// Mitsubishi GX Works2 project: B_v6_split   PLC: Q03UDE

PROGRAM COMMON
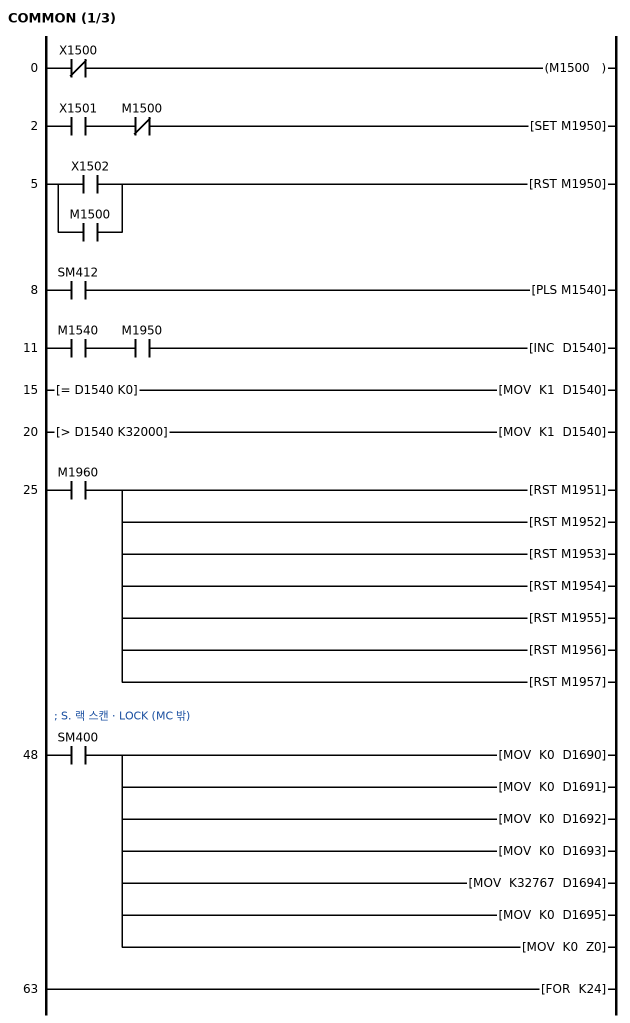
0     LDI     X1500
      OUT     M1500
2     LD      X1501
      ANI     M1500
      SET     M1950
5     LD      X1502
      OR      M1500
      RST     M1950
8     LD      SM412
      PLS     M1540
11    LD      M1540
      AND     M1950
      INC     D1540
15    LD=     D1540 K0
      MOV     K1 D1540
20    LD>     D1540 K32000
      MOV     K1 D1540
25    LD      M1960
      RST     M1951
      RST     M1952
      RST     M1953
      RST     M1954
      RST     M1955
      RST     M1956
      RST     M1957
; S. 랙 스캔 · LOCK (MC 밖)
48    LD      SM400
      MOV     K0 D1690
      MOV     K0 D1691
      MOV     K0 D1692
      MOV     K0 D1693
      MOV     K32767 D1694
      MOV     K0 D1695
      MOV     K0 Z0
63    FOR     K24
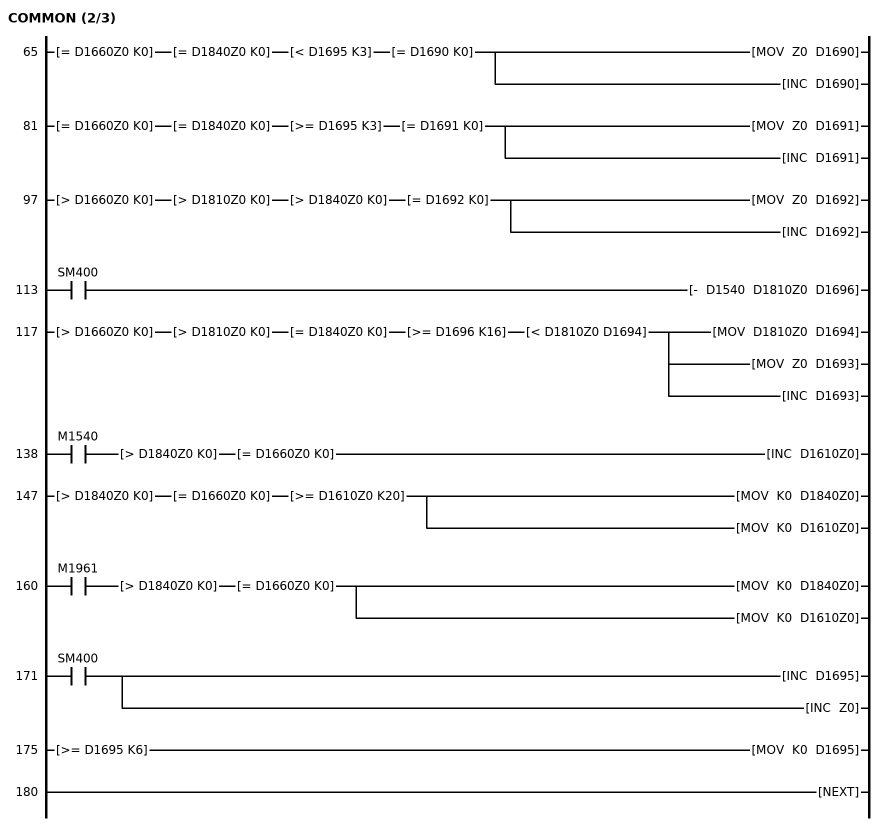
65    LD=     D1660Z0 K0
      AND=    D1840Z0 K0
      AND<    D1695 K3
      AND=    D1690 K0
      MOV     Z0 D1690
      INC     D1690
81    LD=     D1660Z0 K0
      AND=    D1840Z0 K0
      AND>=   D1695 K3
      AND=    D1691 K0
      MOV     Z0 D1691
      INC     D1691
97    LD>     D1660Z0 K0
      AND>    D1810Z0 K0
      AND>    D1840Z0 K0
      AND=    D1692 K0
      MOV     Z0 D1692
      INC     D1692
113   LD      SM400
      -       D1540 D1810Z0 D1696
117   LD>     D1660Z0 K0
      AND>    D1810Z0 K0
      AND=    D1840Z0 K0
      AND>=   D1696 K16
      AND<    D1810Z0 D1694
      MOV     D1810Z0 D1694
      MOV     Z0 D1693
      INC     D1693
138   LD      M1540
      AND>    D1840Z0 K0
      AND=    D1660Z0 K0
      INC     D1610Z0
147   LD>     D1840Z0 K0
      AND=    D1660Z0 K0
      AND>=   D1610Z0 K20
      MOV     K0 D1840Z0
      MOV     K0 D1610Z0
160   LD      M1961
      AND>    D1840Z0 K0
      AND=    D1660Z0 K0
      MOV     K0 D1840Z0
      MOV     K0 D1610Z0
171   LD      SM400
      INC     D1695
      INC     Z0
175   LD>=    D1695 K6
      MOV     K0 D1695
180   NEXT
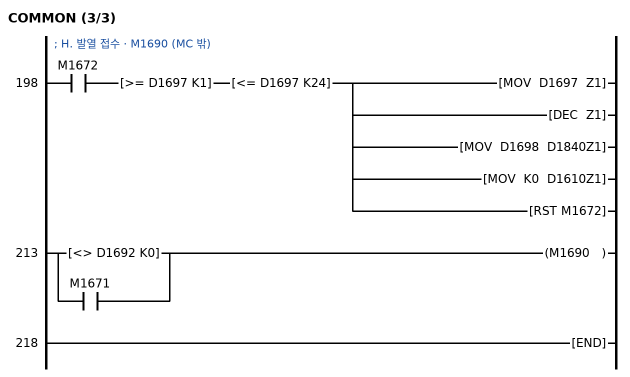
; H. 발열 접수 · M1690 (MC 밖)
198   LD      M1672
      AND>=   D1697 K1
      AND<=   D1697 K24
      MOV     D1697 Z1
      DEC     Z1
      MOV     D1698 D1840Z1
      MOV     K0 D1610Z1
      RST     M1672
213   LD<>    D1692 K0
      OR      M1671
      OUT     M1690
218   END
END_PROGRAM

PROGRAM RFID
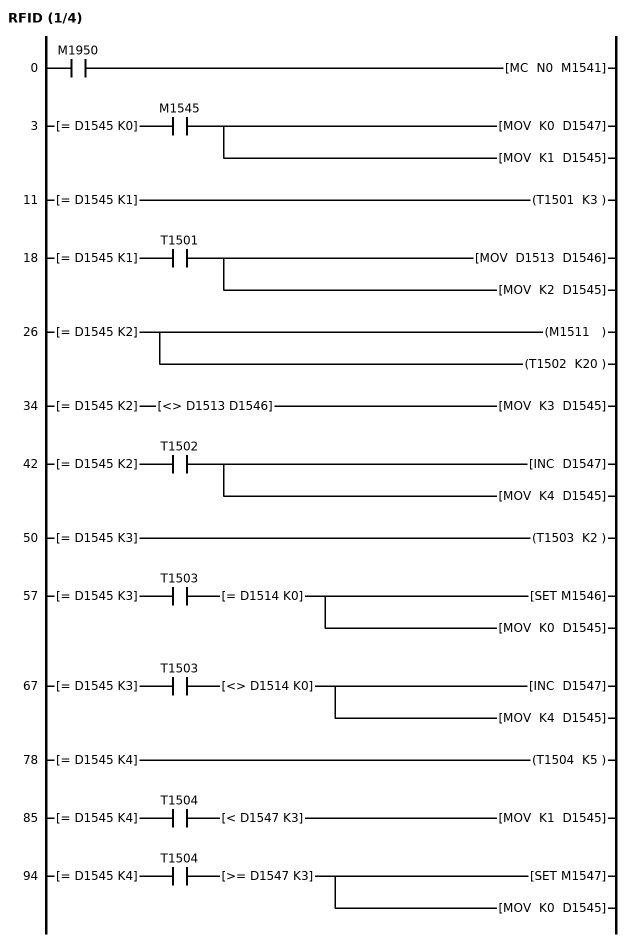
0     LD      M1950
      MC      N0 M1541
3     LD=     D1545 K0
      AND     M1545
      MOV     K0 D1547
      MOV     K1 D1545
11    LD=     D1545 K1
      OUT     T1501 K3
18    LD=     D1545 K1
      AND     T1501
      MOV     D1513 D1546
      MOV     K2 D1545
26    LD=     D1545 K2
      OUT     M1511
      OUT     T1502 K20
34    LD=     D1545 K2
      AND<>   D1513 D1546
      MOV     K3 D1545
42    LD=     D1545 K2
      AND     T1502
      INC     D1547
      MOV     K4 D1545
50    LD=     D1545 K3
      OUT     T1503 K2
57    LD=     D1545 K3
      AND     T1503
      AND=    D1514 K0
      SET     M1546
      MOV     K0 D1545
67    LD=     D1545 K3
      AND     T1503
      AND<>   D1514 K0
      INC     D1547
      MOV     K4 D1545
78    LD=     D1545 K4
      OUT     T1504 K5
85    LD=     D1545 K4
      AND     T1504
      AND<    D1547 K3
      MOV     K1 D1545
94    LD=     D1545 K4
      AND     T1504
      AND>=   D1547 K3
      SET     M1547
      MOV     K0 D1545
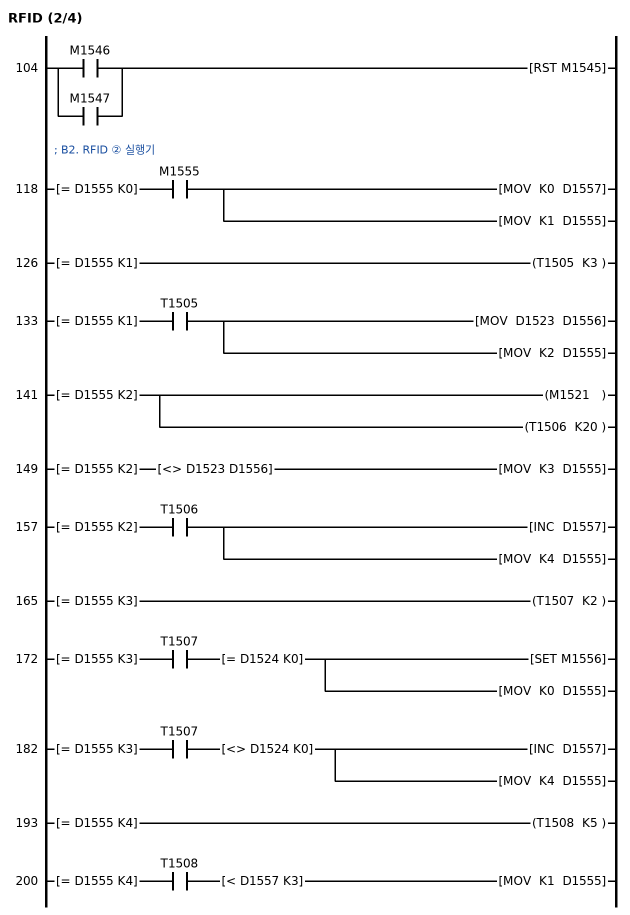
104   LD      M1546
      OR      M1547
      RST     M1545
; B2. RFID ② 실행기
118   LD=     D1555 K0
      AND     M1555
      MOV     K0 D1557
      MOV     K1 D1555
126   LD=     D1555 K1
      OUT     T1505 K3
133   LD=     D1555 K1
      AND     T1505
      MOV     D1523 D1556
      MOV     K2 D1555
141   LD=     D1555 K2
      OUT     M1521
      OUT     T1506 K20
149   LD=     D1555 K2
      AND<>   D1523 D1556
      MOV     K3 D1555
157   LD=     D1555 K2
      AND     T1506
      INC     D1557
      MOV     K4 D1555
165   LD=     D1555 K3
      OUT     T1507 K2
172   LD=     D1555 K3
      AND     T1507
      AND=    D1524 K0
      SET     M1556
      MOV     K0 D1555
182   LD=     D1555 K3
      AND     T1507
      AND<>   D1524 K0
      INC     D1557
      MOV     K4 D1555
193   LD=     D1555 K4
      OUT     T1508 K5
200   LD=     D1555 K4
      AND     T1508
      AND<    D1557 K3
      MOV     K1 D1555
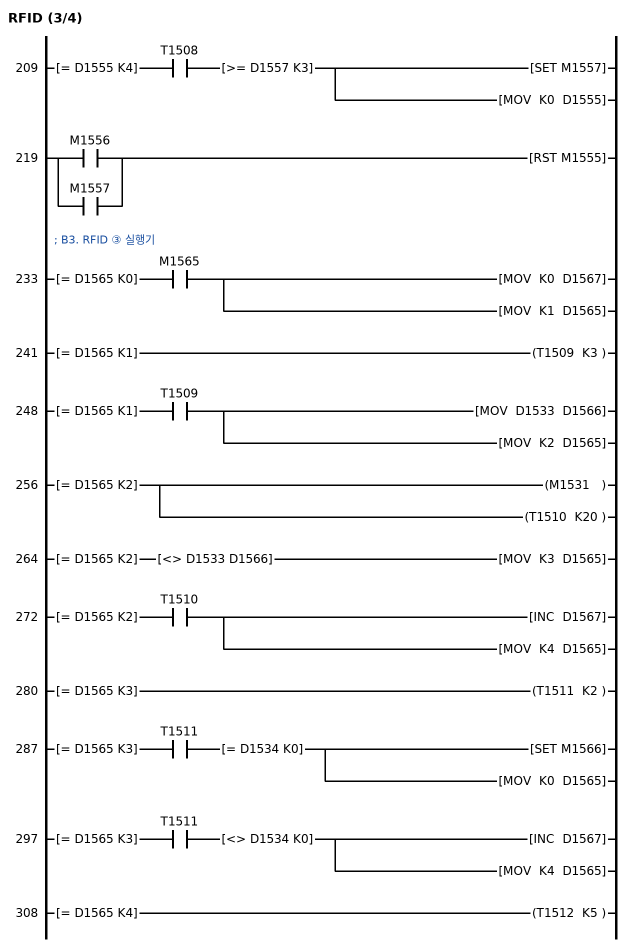
209   LD=     D1555 K4
      AND     T1508
      AND>=   D1557 K3
      SET     M1557
      MOV     K0 D1555
219   LD      M1556
      OR      M1557
      RST     M1555
; B3. RFID ③ 실행기
233   LD=     D1565 K0
      AND     M1565
      MOV     K0 D1567
      MOV     K1 D1565
241   LD=     D1565 K1
      OUT     T1509 K3
248   LD=     D1565 K1
      AND     T1509
      MOV     D1533 D1566
      MOV     K2 D1565
256   LD=     D1565 K2
      OUT     M1531
      OUT     T1510 K20
264   LD=     D1565 K2
      AND<>   D1533 D1566
      MOV     K3 D1565
272   LD=     D1565 K2
      AND     T1510
      INC     D1567
      MOV     K4 D1565
280   LD=     D1565 K3
      OUT     T1511 K2
287   LD=     D1565 K3
      AND     T1511
      AND=    D1534 K0
      SET     M1566
      MOV     K0 D1565
297   LD=     D1565 K3
      AND     T1511
      AND<>   D1534 K0
      INC     D1567
      MOV     K4 D1565
308   LD=     D1565 K4
      OUT     T1512 K5
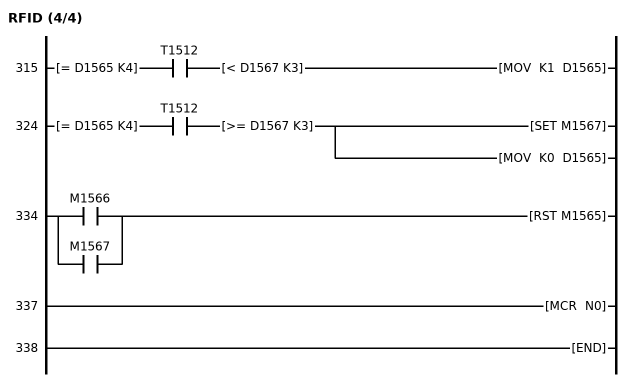
315   LD=     D1565 K4
      AND     T1512
      AND<    D1567 K3
      MOV     K1 D1565
324   LD=     D1565 K4
      AND     T1512
      AND>=   D1567 K3
      SET     M1567
      MOV     K0 D1565
334   LD      M1566
      OR      M1567
      RST     M1565
337   MCR     N0
338   END
END_PROGRAM

PROGRAM INFEED
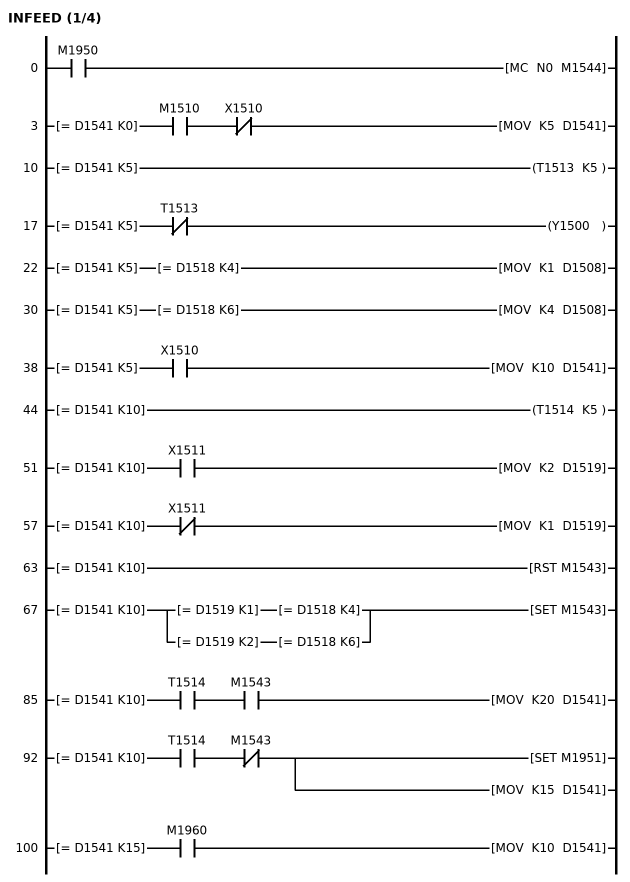
0     LD      M1950
      MC      N0 M1544
3     LD=     D1541 K0
      AND     M1510
      ANI     X1510
      MOV     K5 D1541
10    LD=     D1541 K5
      OUT     T1513 K5
17    LD=     D1541 K5
      ANI     T1513
      OUT     Y1500
22    LD=     D1541 K5
      AND=    D1518 K4
      MOV     K1 D1508
30    LD=     D1541 K5
      AND=    D1518 K6
      MOV     K4 D1508
38    LD=     D1541 K5
      AND     X1510
      MOV     K10 D1541
44    LD=     D1541 K10
      OUT     T1514 K5
51    LD=     D1541 K10
      AND     X1511
      MOV     K2 D1519
57    LD=     D1541 K10
      ANI     X1511
      MOV     K1 D1519
63    LD=     D1541 K10
      RST     M1543
67    LD=     D1541 K10
      LD=     D1519 K1
      AND=    D1518 K4
      LD=     D1519 K2
      AND=    D1518 K6
      ORB
      ANB
      SET     M1543
85    LD=     D1541 K10
      AND     T1514
      AND     M1543
      MOV     K20 D1541
92    LD=     D1541 K10
      AND     T1514
      ANI     M1543
      SET     M1951
      MOV     K15 D1541
100   LD=     D1541 K15
      AND     M1960
      MOV     K10 D1541
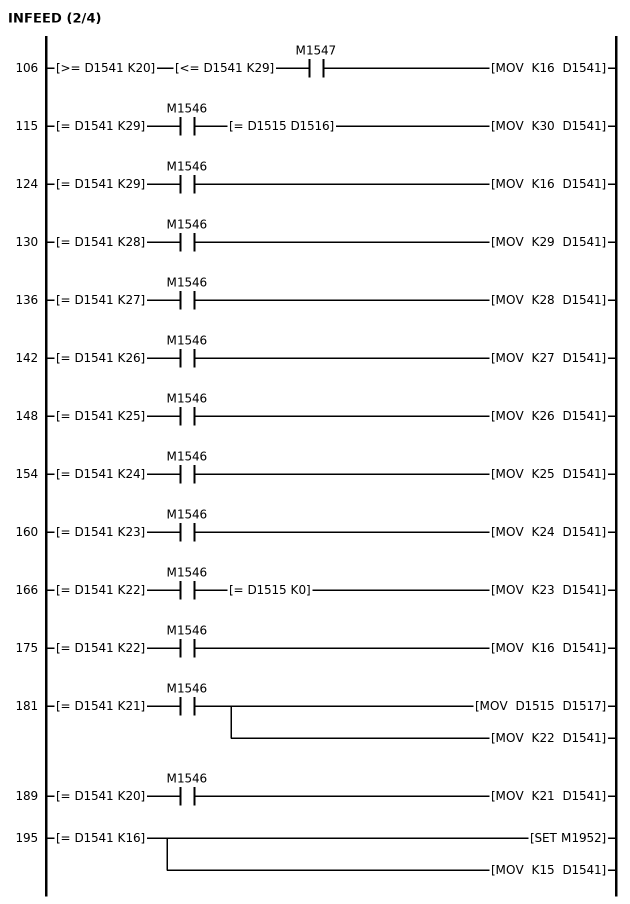
106   LD>=    D1541 K20
      AND<=   D1541 K29
      AND     M1547
      MOV     K16 D1541
115   LD=     D1541 K29
      AND     M1546
      AND=    D1515 D1516
      MOV     K30 D1541
124   LD=     D1541 K29
      AND     M1546
      MOV     K16 D1541
130   LD=     D1541 K28
      AND     M1546
      MOV     K29 D1541
136   LD=     D1541 K27
      AND     M1546
      MOV     K28 D1541
142   LD=     D1541 K26
      AND     M1546
      MOV     K27 D1541
148   LD=     D1541 K25
      AND     M1546
      MOV     K26 D1541
154   LD=     D1541 K24
      AND     M1546
      MOV     K25 D1541
160   LD=     D1541 K23
      AND     M1546
      MOV     K24 D1541
166   LD=     D1541 K22
      AND     M1546
      AND=    D1515 K0
      MOV     K23 D1541
175   LD=     D1541 K22
      AND     M1546
      MOV     K16 D1541
181   LD=     D1541 K21
      AND     M1546
      MOV     D1515 D1517
      MOV     K22 D1541
189   LD=     D1541 K20
      AND     M1546
      MOV     K21 D1541
195   LD=     D1541 K16
      SET     M1952
      MOV     K15 D1541
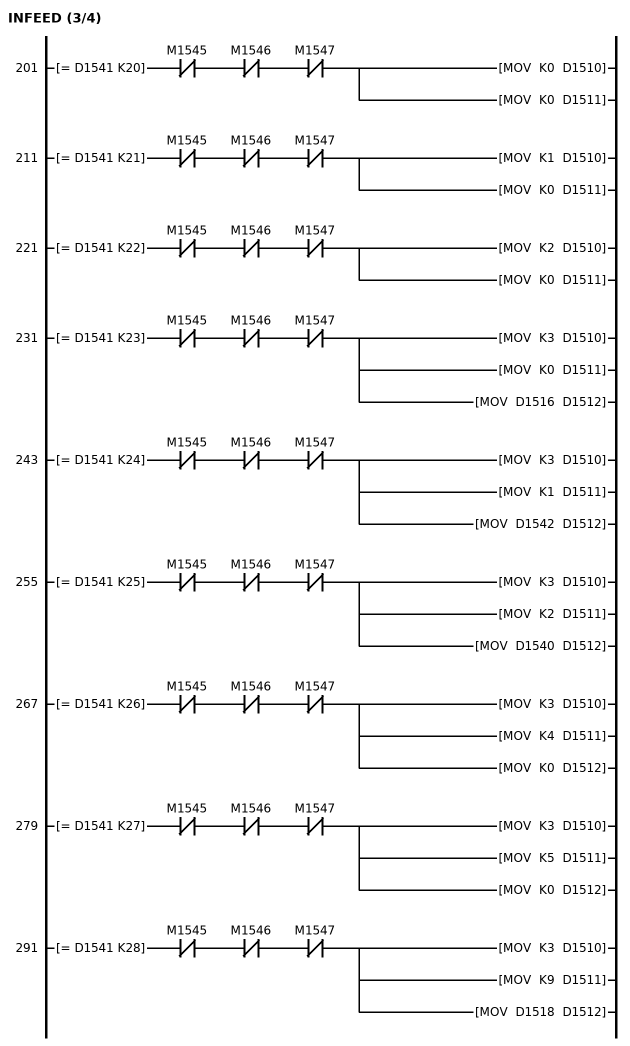
201   LD=     D1541 K20
      ANI     M1545
      ANI     M1546
      ANI     M1547
      MOV     K0 D1510
      MOV     K0 D1511
211   LD=     D1541 K21
      ANI     M1545
      ANI     M1546
      ANI     M1547
      MOV     K1 D1510
      MOV     K0 D1511
221   LD=     D1541 K22
      ANI     M1545
      ANI     M1546
      ANI     M1547
      MOV     K2 D1510
      MOV     K0 D1511
231   LD=     D1541 K23
      ANI     M1545
      ANI     M1546
      ANI     M1547
      MOV     K3 D1510
      MOV     K0 D1511
      MOV     D1516 D1512
243   LD=     D1541 K24
      ANI     M1545
      ANI     M1546
      ANI     M1547
      MOV     K3 D1510
      MOV     K1 D1511
      MOV     D1542 D1512
255   LD=     D1541 K25
      ANI     M1545
      ANI     M1546
      ANI     M1547
      MOV     K3 D1510
      MOV     K2 D1511
      MOV     D1540 D1512
267   LD=     D1541 K26
      ANI     M1545
      ANI     M1546
      ANI     M1547
      MOV     K3 D1510
      MOV     K4 D1511
      MOV     K0 D1512
279   LD=     D1541 K27
      ANI     M1545
      ANI     M1546
      ANI     M1547
      MOV     K3 D1510
      MOV     K5 D1511
      MOV     K0 D1512
291   LD=     D1541 K28
      ANI     M1545
      ANI     M1546
      ANI     M1547
      MOV     K3 D1510
      MOV     K9 D1511
      MOV     D1518 D1512
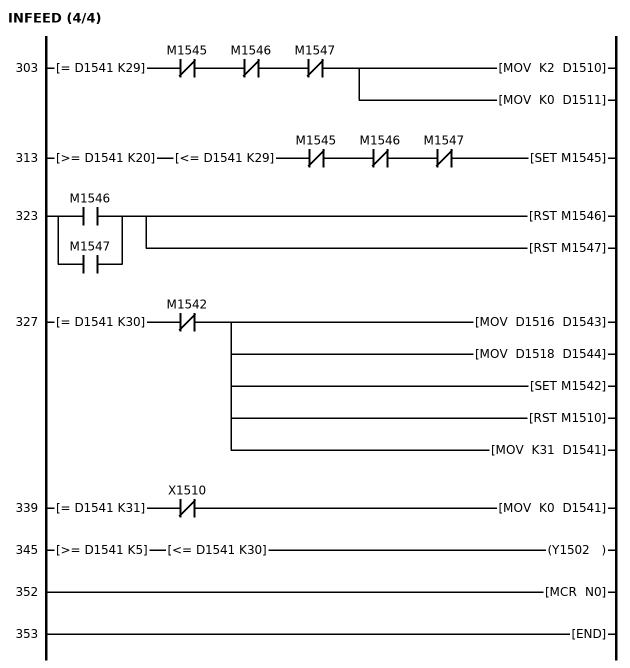
303   LD=     D1541 K29
      ANI     M1545
      ANI     M1546
      ANI     M1547
      MOV     K2 D1510
      MOV     K0 D1511
313   LD>=    D1541 K20
      AND<=   D1541 K29
      ANI     M1545
      ANI     M1546
      ANI     M1547
      SET     M1545
323   LD      M1546
      OR      M1547
      RST     M1546
      RST     M1547
327   LD=     D1541 K30
      ANI     M1542
      MOV     D1516 D1543
      MOV     D1518 D1544
      SET     M1542
      RST     M1510
      MOV     K31 D1541
339   LD=     D1541 K31
      ANI     X1510
      MOV     K0 D1541
345   LD>=    D1541 K5
      AND<=   D1541 K30
      OUT     Y1502
352   MCR     N0
353   END
END_PROGRAM

PROGRAM CRANE
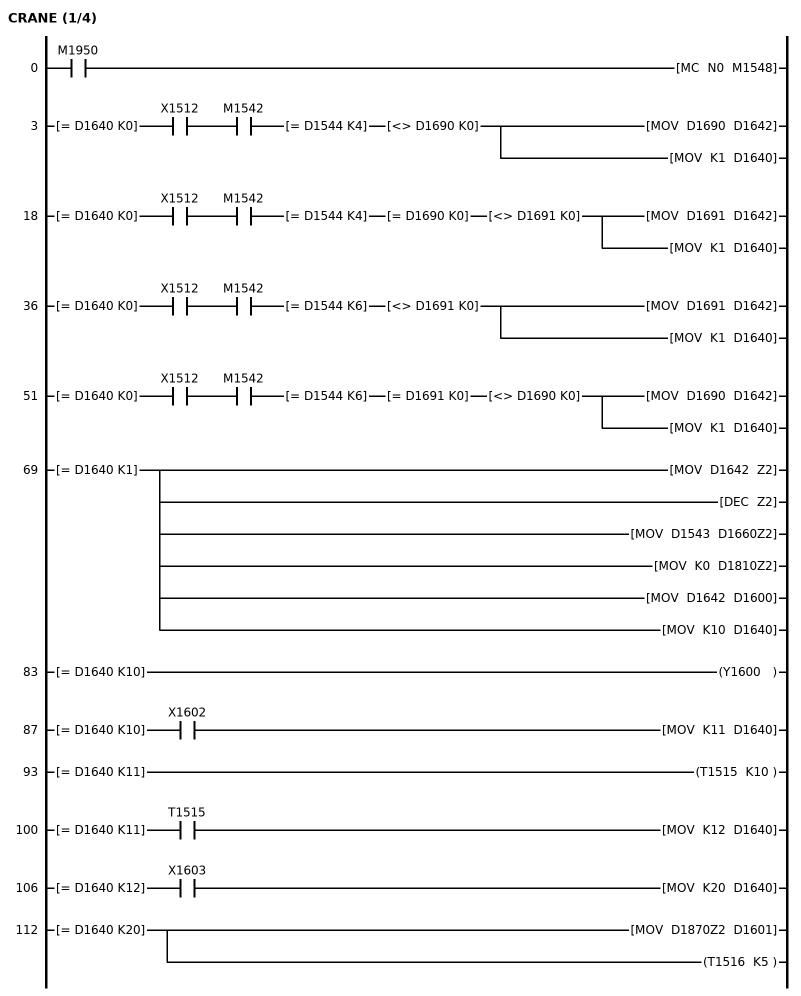
0     LD      M1950
      MC      N0 M1548
3     LD=     D1640 K0
      AND     X1512
      AND     M1542
      AND=    D1544 K4
      AND<>   D1690 K0
      MOV     D1690 D1642
      MOV     K1 D1640
18    LD=     D1640 K0
      AND     X1512
      AND     M1542
      AND=    D1544 K4
      AND=    D1690 K0
      AND<>   D1691 K0
      MOV     D1691 D1642
      MOV     K1 D1640
36    LD=     D1640 K0
      AND     X1512
      AND     M1542
      AND=    D1544 K6
      AND<>   D1691 K0
      MOV     D1691 D1642
      MOV     K1 D1640
51    LD=     D1640 K0
      AND     X1512
      AND     M1542
      AND=    D1544 K6
      AND=    D1691 K0
      AND<>   D1690 K0
      MOV     D1690 D1642
      MOV     K1 D1640
69    LD=     D1640 K1
      MOV     D1642 Z2
      DEC     Z2
      MOV     D1543 D1660Z2
      MOV     K0 D1810Z2
      MOV     D1642 D1600
      MOV     K10 D1640
83    LD=     D1640 K10
      OUT     Y1600
87    LD=     D1640 K10
      AND     X1602
      MOV     K11 D1640
93    LD=     D1640 K11
      OUT     T1515 K10
100   LD=     D1640 K11
      AND     T1515
      MOV     K12 D1640
106   LD=     D1640 K12
      AND     X1603
      MOV     K20 D1640
112   LD=     D1640 K20
      MOV     D1870Z2 D1601
      OUT     T1516 K5
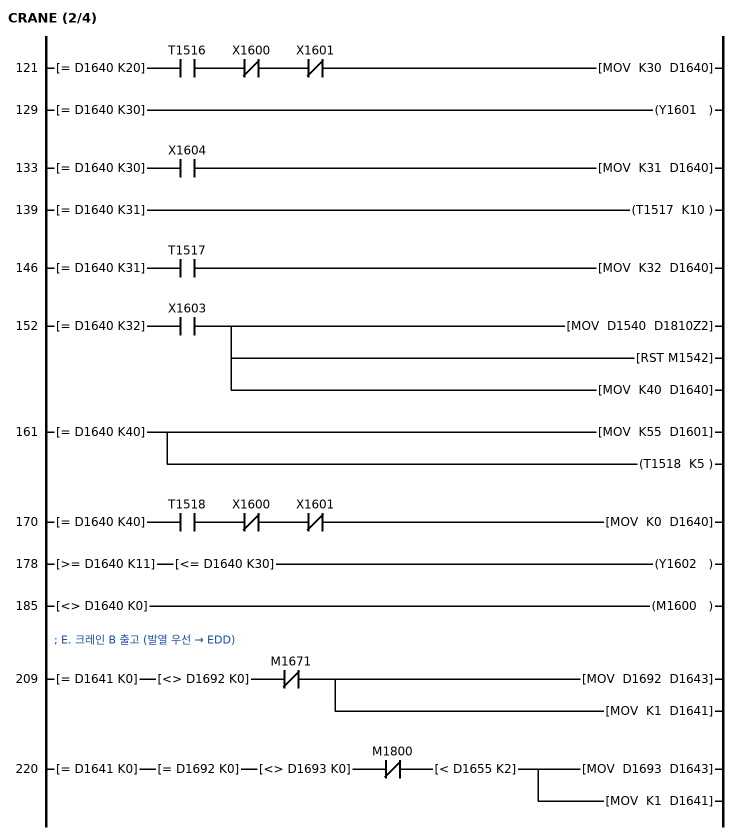
121   LD=     D1640 K20
      AND     T1516
      ANI     X1600
      ANI     X1601
      MOV     K30 D1640
129   LD=     D1640 K30
      OUT     Y1601
133   LD=     D1640 K30
      AND     X1604
      MOV     K31 D1640
139   LD=     D1640 K31
      OUT     T1517 K10
146   LD=     D1640 K31
      AND     T1517
      MOV     K32 D1640
152   LD=     D1640 K32
      AND     X1603
      MOV     D1540 D1810Z2
      RST     M1542
      MOV     K40 D1640
161   LD=     D1640 K40
      MOV     K55 D1601
      OUT     T1518 K5
170   LD=     D1640 K40
      AND     T1518
      ANI     X1600
      ANI     X1601
      MOV     K0 D1640
178   LD>=    D1640 K11
      AND<=   D1640 K30
      OUT     Y1602
185   LD<>    D1640 K0
      OUT     M1600
; E. 크레인 B 출고 (발열 우선 → EDD)
209   LD=     D1641 K0
      AND<>   D1692 K0
      ANI     M1671
      MOV     D1692 D1643
      MOV     K1 D1641
220   LD=     D1641 K0
      AND=    D1692 K0
      AND<>   D1693 K0
      ANI     M1800
      AND<    D1655 K2
      MOV     D1693 D1643
      MOV     K1 D1641
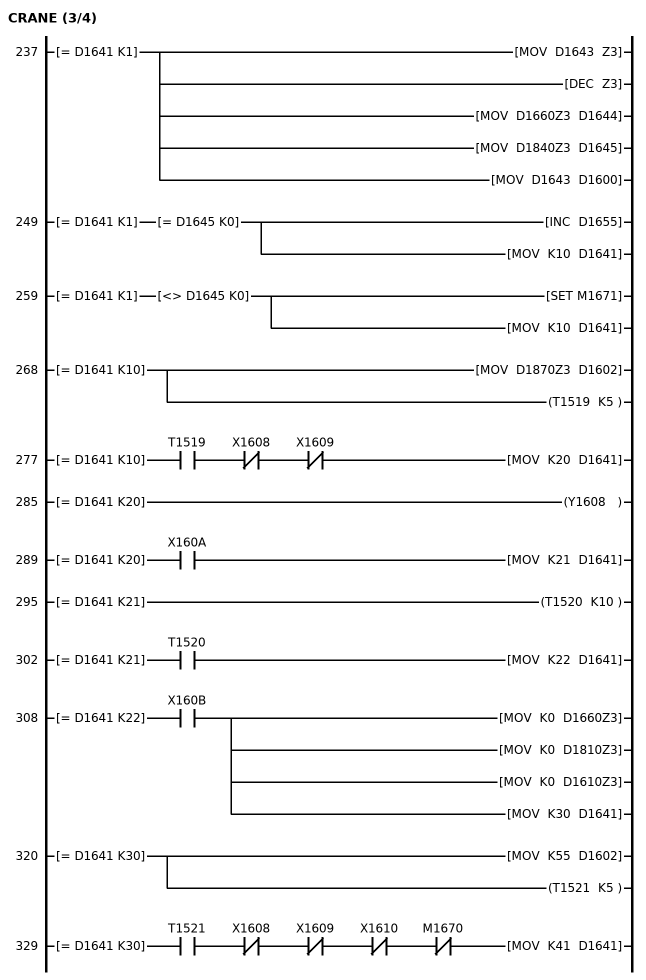
237   LD=     D1641 K1
      MOV     D1643 Z3
      DEC     Z3
      MOV     D1660Z3 D1644
      MOV     D1840Z3 D1645
      MOV     D1643 D1600
249   LD=     D1641 K1
      AND=    D1645 K0
      INC     D1655
      MOV     K10 D1641
259   LD=     D1641 K1
      AND<>   D1645 K0
      SET     M1671
      MOV     K10 D1641
268   LD=     D1641 K10
      MOV     D1870Z3 D1602
      OUT     T1519 K5
277   LD=     D1641 K10
      AND     T1519
      ANI     X1608
      ANI     X1609
      MOV     K20 D1641
285   LD=     D1641 K20
      OUT     Y1608
289   LD=     D1641 K20
      AND     X160A
      MOV     K21 D1641
295   LD=     D1641 K21
      OUT     T1520 K10
302   LD=     D1641 K21
      AND     T1520
      MOV     K22 D1641
308   LD=     D1641 K22
      AND     X160B
      MOV     K0 D1660Z3
      MOV     K0 D1810Z3
      MOV     K0 D1610Z3
      MOV     K30 D1641
320   LD=     D1641 K30
      MOV     K55 D1602
      OUT     T1521 K5
329   LD=     D1641 K30
      AND     T1521
      ANI     X1608
      ANI     X1609
      ANI     X1610
      ANI     M1670
      MOV     K41 D1641
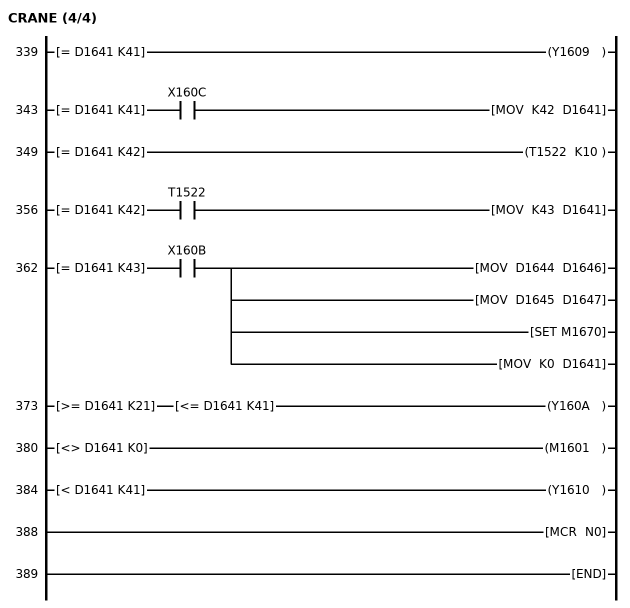
339   LD=     D1641 K41
      OUT     Y1609
343   LD=     D1641 K41
      AND     X160C
      MOV     K42 D1641
349   LD=     D1641 K42
      OUT     T1522 K10
356   LD=     D1641 K42
      AND     T1522
      MOV     K43 D1641
362   LD=     D1641 K43
      AND     X160B
      MOV     D1644 D1646
      MOV     D1645 D1647
      SET     M1670
      MOV     K0 D1641
373   LD>=    D1641 K21
      AND<=   D1641 K41
      OUT     Y160A
380   LD<>    D1641 K0
      OUT     M1601
384   LD<     D1641 K41
      OUT     Y1610
388   MCR     N0
389   END
END_PROGRAM

PROGRAM SORT1
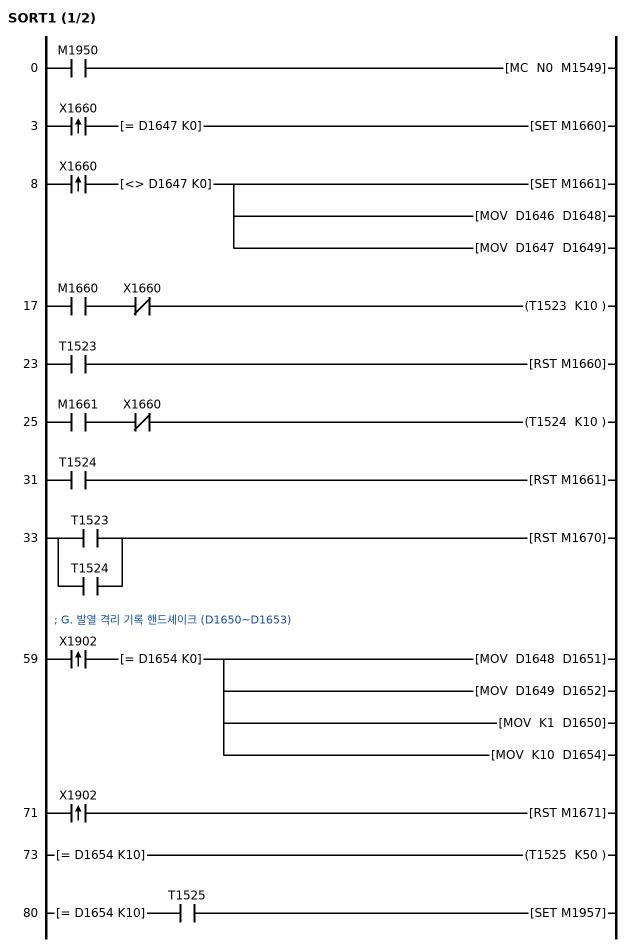
0     LD      M1950
      MC      N0 M1549
3     LDP     X1660
      AND=    D1647 K0
      SET     M1660
8     LDP     X1660
      AND<>   D1647 K0
      SET     M1661
      MOV     D1646 D1648
      MOV     D1647 D1649
17    LD      M1660
      ANI     X1660
      OUT     T1523 K10
23    LD      T1523
      RST     M1660
25    LD      M1661
      ANI     X1660
      OUT     T1524 K10
31    LD      T1524
      RST     M1661
33    LD      T1523
      OR      T1524
      RST     M1670
; G. 발열 격리 기록 핸드셰이크 (D1650~D1653)
59    LDP     X1902
      AND=    D1654 K0
      MOV     D1648 D1651
      MOV     D1649 D1652
      MOV     K1 D1650
      MOV     K10 D1654
71    LDP     X1902
      RST     M1671
73    LD=     D1654 K10
      OUT     T1525 K50
80    LD=     D1654 K10
      AND     T1525
      SET     M1957
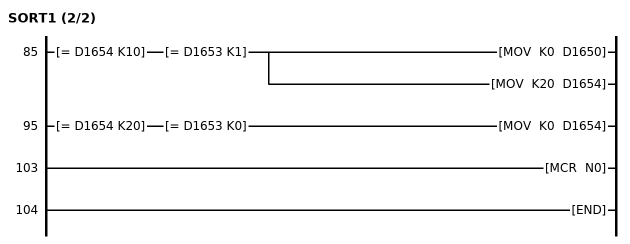
85    LD=     D1654 K10
      AND=    D1653 K1
      MOV     K0 D1650
      MOV     K20 D1654
95    LD=     D1654 K20
      AND=    D1653 K0
      MOV     K0 D1654
103   MCR     N0
104   END
END_PROGRAM

PROGRAM INSPECT
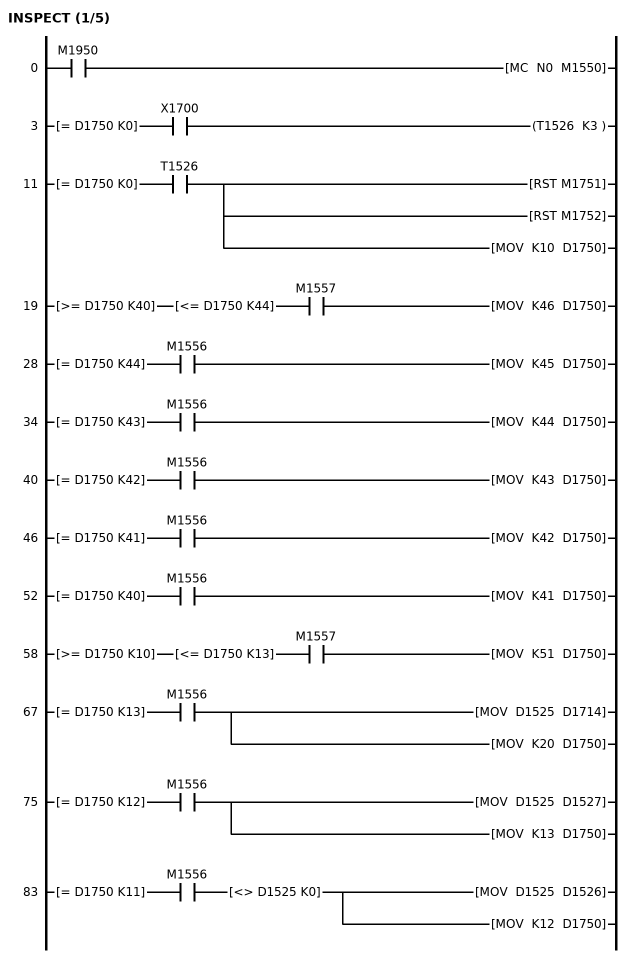
0     LD      M1950
      MC      N0 M1550
3     LD=     D1750 K0
      AND     X1700
      OUT     T1526 K3
11    LD=     D1750 K0
      AND     T1526
      RST     M1751
      RST     M1752
      MOV     K10 D1750
19    LD>=    D1750 K40
      AND<=   D1750 K44
      AND     M1557
      MOV     K46 D1750
28    LD=     D1750 K44
      AND     M1556
      MOV     K45 D1750
34    LD=     D1750 K43
      AND     M1556
      MOV     K44 D1750
40    LD=     D1750 K42
      AND     M1556
      MOV     K43 D1750
46    LD=     D1750 K41
      AND     M1556
      MOV     K42 D1750
52    LD=     D1750 K40
      AND     M1556
      MOV     K41 D1750
58    LD>=    D1750 K10
      AND<=   D1750 K13
      AND     M1557
      MOV     K51 D1750
67    LD=     D1750 K13
      AND     M1556
      MOV     D1525 D1714
      MOV     K20 D1750
75    LD=     D1750 K12
      AND     M1556
      MOV     D1525 D1527
      MOV     K13 D1750
83    LD=     D1750 K11
      AND     M1556
      AND<>   D1525 K0
      MOV     D1525 D1526
      MOV     K12 D1750
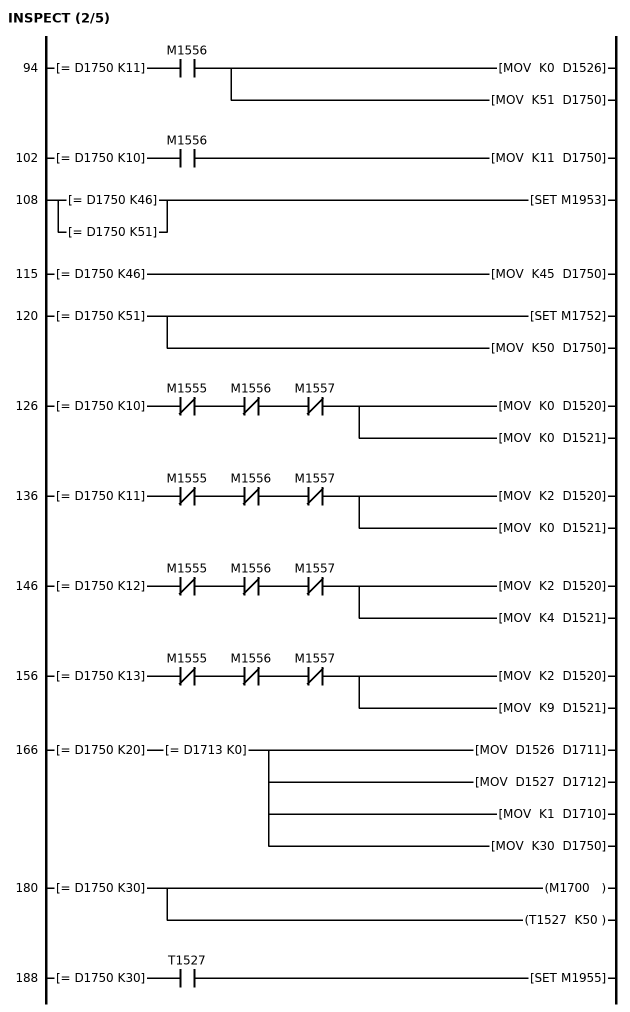
94    LD=     D1750 K11
      AND     M1556
      MOV     K0 D1526
      MOV     K51 D1750
102   LD=     D1750 K10
      AND     M1556
      MOV     K11 D1750
108   LD=     D1750 K46
      OR=     D1750 K51
      SET     M1953
115   LD=     D1750 K46
      MOV     K45 D1750
120   LD=     D1750 K51
      SET     M1752
      MOV     K50 D1750
126   LD=     D1750 K10
      ANI     M1555
      ANI     M1556
      ANI     M1557
      MOV     K0 D1520
      MOV     K0 D1521
136   LD=     D1750 K11
      ANI     M1555
      ANI     M1556
      ANI     M1557
      MOV     K2 D1520
      MOV     K0 D1521
146   LD=     D1750 K12
      ANI     M1555
      ANI     M1556
      ANI     M1557
      MOV     K2 D1520
      MOV     K4 D1521
156   LD=     D1750 K13
      ANI     M1555
      ANI     M1556
      ANI     M1557
      MOV     K2 D1520
      MOV     K9 D1521
166   LD=     D1750 K20
      AND=    D1713 K0
      MOV     D1526 D1711
      MOV     D1527 D1712
      MOV     K1 D1710
      MOV     K30 D1750
180   LD=     D1750 K30
      OUT     M1700
      OUT     T1527 K50
188   LD=     D1750 K30
      AND     T1527
      SET     M1955
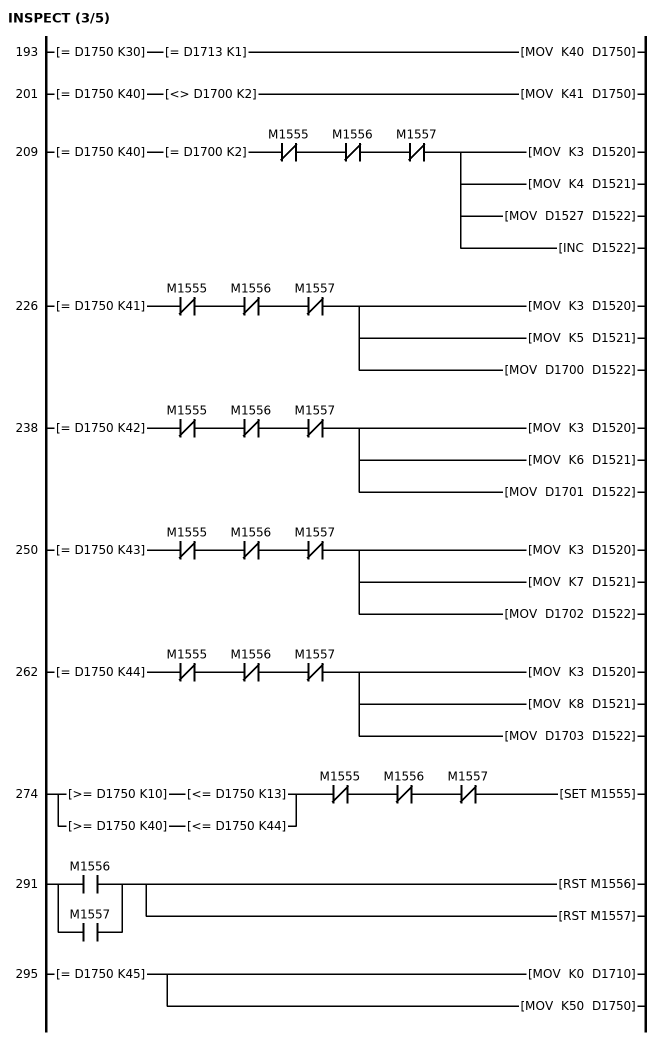
193   LD=     D1750 K30
      AND=    D1713 K1
      MOV     K40 D1750
201   LD=     D1750 K40
      AND<>   D1700 K2
      MOV     K41 D1750
209   LD=     D1750 K40
      AND=    D1700 K2
      ANI     M1555
      ANI     M1556
      ANI     M1557
      MOV     K3 D1520
      MOV     K4 D1521
      MOV     D1527 D1522
      INC     D1522
226   LD=     D1750 K41
      ANI     M1555
      ANI     M1556
      ANI     M1557
      MOV     K3 D1520
      MOV     K5 D1521
      MOV     D1700 D1522
238   LD=     D1750 K42
      ANI     M1555
      ANI     M1556
      ANI     M1557
      MOV     K3 D1520
      MOV     K6 D1521
      MOV     D1701 D1522
250   LD=     D1750 K43
      ANI     M1555
      ANI     M1556
      ANI     M1557
      MOV     K3 D1520
      MOV     K7 D1521
      MOV     D1702 D1522
262   LD=     D1750 K44
      ANI     M1555
      ANI     M1556
      ANI     M1557
      MOV     K3 D1520
      MOV     K8 D1521
      MOV     D1703 D1522
274   LD>=    D1750 K10
      AND<=   D1750 K13
      LD>=    D1750 K40
      AND<=   D1750 K44
      ORB
      ANI     M1555
      ANI     M1556
      ANI     M1557
      SET     M1555
291   LD      M1556
      OR      M1557
      RST     M1556
      RST     M1557
295   LD=     D1750 K45
      MOV     K0 D1710
      MOV     K50 D1750
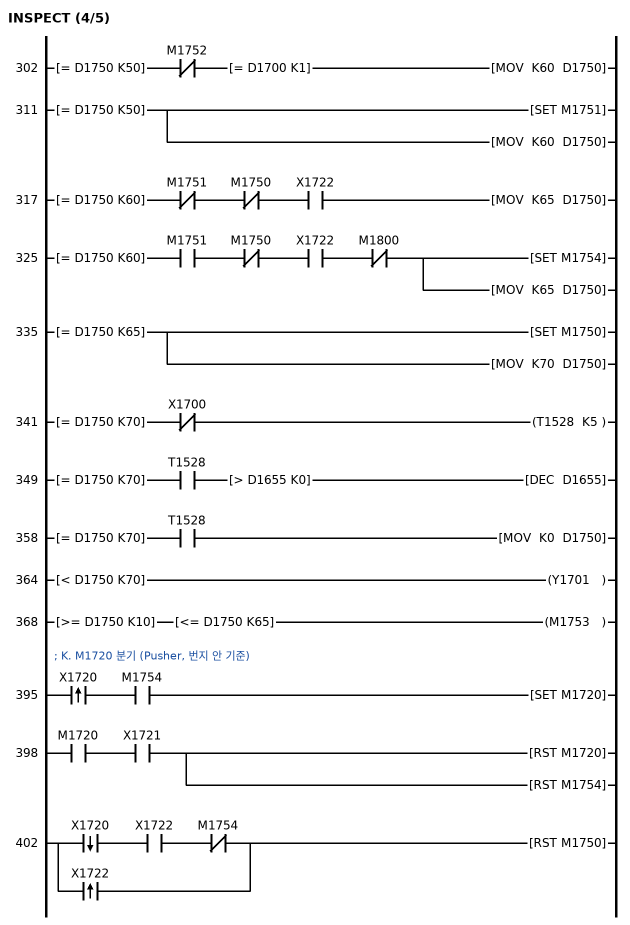
302   LD=     D1750 K50
      ANI     M1752
      AND=    D1700 K1
      MOV     K60 D1750
311   LD=     D1750 K50
      SET     M1751
      MOV     K60 D1750
317   LD=     D1750 K60
      ANI     M1751
      ANI     M1750
      AND     X1722
      MOV     K65 D1750
325   LD=     D1750 K60
      AND     M1751
      ANI     M1750
      AND     X1722
      ANI     M1800
      SET     M1754
      MOV     K65 D1750
335   LD=     D1750 K65
      SET     M1750
      MOV     K70 D1750
341   LD=     D1750 K70
      ANI     X1700
      OUT     T1528 K5
349   LD=     D1750 K70
      AND     T1528
      AND>    D1655 K0
      DEC     D1655
358   LD=     D1750 K70
      AND     T1528
      MOV     K0 D1750
364   LD<     D1750 K70
      OUT     Y1701
368   LD>=    D1750 K10
      AND<=   D1750 K65
      OUT     M1753
; K. M1720 분기 (Pusher, 번지 안 기준)
395   LDP     X1720
      AND     M1754
      SET     M1720
398   LD      M1720
      AND     X1721
      RST     M1720
      RST     M1754
402   LDF     X1720
      AND     X1722
      ANI     M1754
      ORP     X1722
      RST     M1750
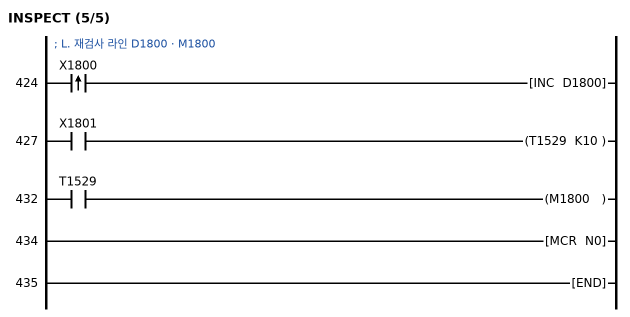
; L. 재검사 라인 D1800 · M1800
424   LDP     X1800
      INC     D1800
427   LD      X1801
      OUT     T1529 K10
432   LD      T1529
      OUT     M1800
434   MCR     N0
435   END
END_PROGRAM

PROGRAM RETEST
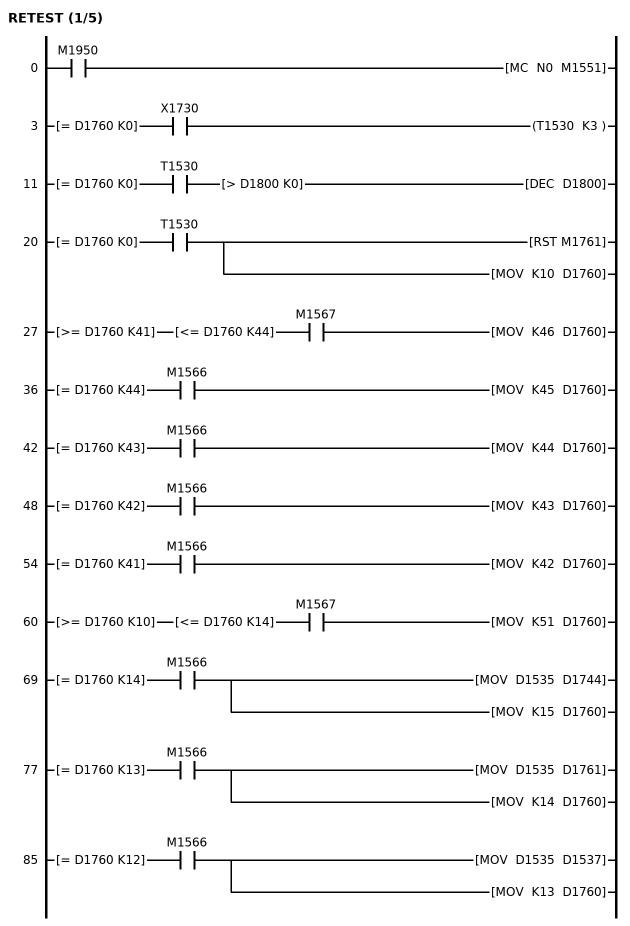
0     LD      M1950
      MC      N0 M1551
3     LD=     D1760 K0
      AND     X1730
      OUT     T1530 K3
11    LD=     D1760 K0
      AND     T1530
      AND>    D1800 K0
      DEC     D1800
20    LD=     D1760 K0
      AND     T1530
      RST     M1761
      MOV     K10 D1760
27    LD>=    D1760 K41
      AND<=   D1760 K44
      AND     M1567
      MOV     K46 D1760
36    LD=     D1760 K44
      AND     M1566
      MOV     K45 D1760
42    LD=     D1760 K43
      AND     M1566
      MOV     K44 D1760
48    LD=     D1760 K42
      AND     M1566
      MOV     K43 D1760
54    LD=     D1760 K41
      AND     M1566
      MOV     K42 D1760
60    LD>=    D1760 K10
      AND<=   D1760 K14
      AND     M1567
      MOV     K51 D1760
69    LD=     D1760 K14
      AND     M1566
      MOV     D1535 D1744
      MOV     K15 D1760
77    LD=     D1760 K13
      AND     M1566
      MOV     D1535 D1761
      MOV     K14 D1760
85    LD=     D1760 K12
      AND     M1566
      MOV     D1535 D1537
      MOV     K13 D1760
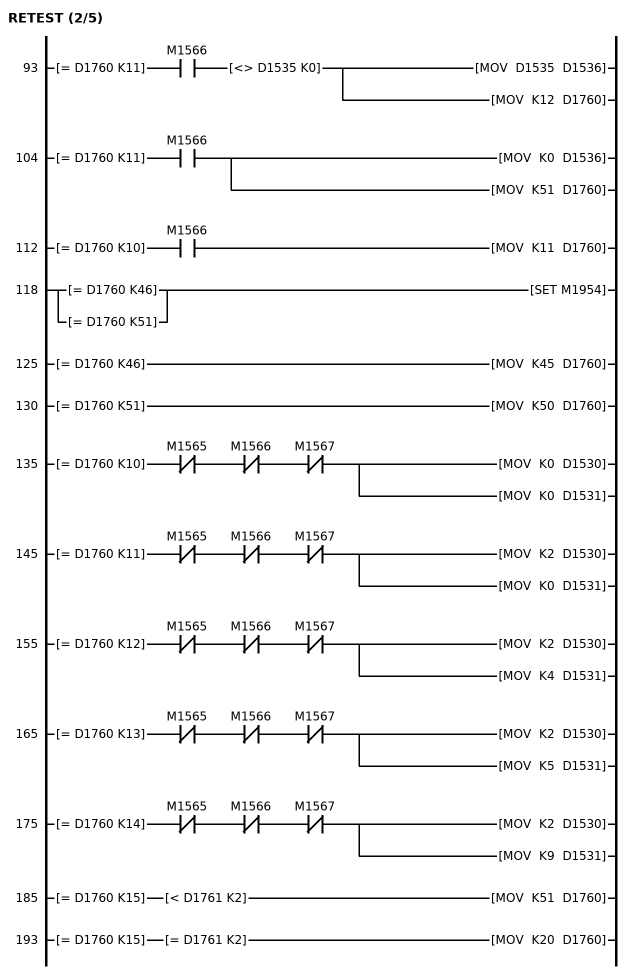
93    LD=     D1760 K11
      AND     M1566
      AND<>   D1535 K0
      MOV     D1535 D1536
      MOV     K12 D1760
104   LD=     D1760 K11
      AND     M1566
      MOV     K0 D1536
      MOV     K51 D1760
112   LD=     D1760 K10
      AND     M1566
      MOV     K11 D1760
118   LD=     D1760 K46
      OR=     D1760 K51
      SET     M1954
125   LD=     D1760 K46
      MOV     K45 D1760
130   LD=     D1760 K51
      MOV     K50 D1760
135   LD=     D1760 K10
      ANI     M1565
      ANI     M1566
      ANI     M1567
      MOV     K0 D1530
      MOV     K0 D1531
145   LD=     D1760 K11
      ANI     M1565
      ANI     M1566
      ANI     M1567
      MOV     K2 D1530
      MOV     K0 D1531
155   LD=     D1760 K12
      ANI     M1565
      ANI     M1566
      ANI     M1567
      MOV     K2 D1530
      MOV     K4 D1531
165   LD=     D1760 K13
      ANI     M1565
      ANI     M1566
      ANI     M1567
      MOV     K2 D1530
      MOV     K5 D1531
175   LD=     D1760 K14
      ANI     M1565
      ANI     M1566
      ANI     M1567
      MOV     K2 D1530
      MOV     K9 D1531
185   LD=     D1760 K15
      AND<    D1761 K2
      MOV     K51 D1760
193   LD=     D1760 K15
      AND=    D1761 K2
      MOV     K20 D1760
